Fanuc KAREL source: KT00628.KL

PROGRAM KT00628
%NOLOCKGROUP
VAR
  S1: STRING[80]
  S2: STRING[80]
  OUT: INTEGER
BEGIN
  S1 = 'A'
  S2 = 'B'
  S1 = 'A'
  S2 = 'B'
  OUT = + S1
END KT00628
